// TIA Portal V21 export
// export: Created 2026-11-21T13:31:41.8064337Z, ExportSetting WithDefaults, DisplayName Totally Integrated Automation Portal, DisplayVersion V21, DisplayName STEP 7 Professional, DisplayVersion V21, DisplayName STEP 7 Safety, DisplayVersion V21, DisplayName Tech WebApplication, DisplayVersion V21, DisplayName WinCC Basic/Comfort/Advanced, DisplayVersion V21, DisplayName WinCC Unified, DisplayVersion V21
FUNCTION_BLOCK "Timed"   // FB30, GRAPH
TITLE = Timed carriage
VERSION : 0.1
// A carriage that runs and brakes, with step times: the defaults, both set, and only the maximum set.
// stored: AcknowledgeErrorsRequired true, AutoNumber true, GraphVersion 6.0, InitialValuesAcquisition false, IsIECCheckEnabled false, LanguageInNetworks LAD, LockOperatingMode false, PermanentILProcessingInMANMode false, SetENOAutomatically false, SkipSteps false, UDAEnableTagReadback false, WithAlarmHandling true
   // inherited from GRAPH_BASE
   VAR
      OFF_SQ_BASE : Bool;
   END_VAR
   VAR_INPUT
      ACK_EF : Bool := false;   // Acknowledge all errors and faults
      go : Bool;
      arrived : Bool;
      stopped : Bool;
      jammed : Bool;
   END_VAR
   VAR_OUTPUT
      motor : Bool;
      brake : Bool;
   END_VAR
BEGIN
// Sequence
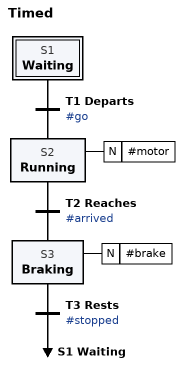
   // sequencer 1
   INITIAL_STEP Waiting:   // S1, max time T#10S, warning time T#7S
   END_STEP
   TRANSITION Departs FROM Waiting TO Running   // T1
      := #go;
   END_TRANSITION
   STEP Running:   // S2, max time T#30S, warning time T#20S
      supervision V := #jammed;
              N    #motor
   END_STEP
   TRANSITION Reaches FROM Running TO Braking   // T2
      := #arrived;
   END_TRANSITION
   STEP Braking:   // S3, max time T#1M30S, warning time T#7S
              N    #brake
   END_STEP
   TRANSITION Rests FROM Braking TO Waiting   // T3, jump
      := #stopped;
   END_TRANSITION
END_FUNCTION_BLOCK
